Fanuc KAREL source: KT00892.KL

PROGRAM KT00892
%NOLOCKGROUP
VAR
  V1: VECTOR
  V2: VECTOR
  OUT: POSITION
BEGIN
  V1.X = 1.0
  V2.Y = 2.0
  V1.X = 1.0
  V2.Y = 2.0
  OUT = INV(V1)
END KT00892
